(*
SPDX-FileCopyrightText: © 2026 Oleksandr Tiutyk <trofimich@gmail.com>
SPDX-License-Identifier: MIT
License: https://opensource.org/license/mit
*)

(*!
<summary>
Defines the contract for an activity that executes an asynchronous task from TwinCAT.OpenFramework.Tasks.
</summary>
<description>
Starts the task on entry, cyclically executes it while RUNNING, translates stop reasons (WORK_DONE to
completion, INTERNAL_ABORT or EXTERNAL_CANCEL to halted, FAILURE to exception) and propagates cancellation
requests to the task. While suspending, the task keeps executing until it stops. A task failure during
stopping is still an activity failure; work completion completes the activity rather than reporting a pause.
Persistent task bindings distinguish a workflow-owned configuration from an external key.
</description>
*)

INTERFACE IInvokeTaskActivity EXTENDS IActivity

(*!
<summary>Reports whether the task activity has been configured.</summary>
*)
{attribute 'monitoring' := 'call'}
PROPERTY Configured : BOOL
GET
END_GET
END_PROPERTY

(*!
<summary>Configures the task to be executed.</summary>
<description>
Requires a nonzero task instance and PASSIVE_READY. The task is borrowed until stopping and reset finish.
This execution-only binding clears any previously configured persistence role.
Rejected configuration preserves the previous dependency; active task replacement is not supported.
</description>
<param name="task">The task instance to execute.</param>
*)
METHOD Configure
VAR_INPUT
	task : TOF_Tasks.ITask;
END_VAR
END_METHOD

(*!
<summary>Returns the configured task instance, or 0 before configuration.</summary>
*)
{attribute 'monitoring' := 'call'}
PROPERTY Task : TOF_Tasks.ITask
GET
END_GET
END_PROPERTY

(*!
<summary>Adopts a fresh workflow-owned task.</summary>
<description>Requires a ready node in a workflow and a dynamic serializable instance available for exclusive transfer.
The workflow owns it on success. A duplicate in the same workflow raises before changing this node.</description>
*)
METHOD ConfigureEmbeddedTask
VAR_INPUT
	task : TOF_Tasks.ITask;
END_VAR
END_METHOD

(*!
<summary>Binds an externally owned task.</summary>
<description>Requires a live dependency and a nonempty stable key. Several nodes may borrow the same external instance.
The provider keeps it alive. Rejection preserves the previous binding.</description>
*)
METHOD ConfigureExternalTask
VAR_INPUT
	task : TOF_Tasks.ITask;
	key : STRING;
END_VAR
END_METHOD

END_INTERFACE

(* stored: Version 1.1.0.1
   Itf IInvokeTaskActivity: Id {4aac828c-d9ae-42b7-9869-9d06d2ade0db}
   Property Configured: Id {63c9557d-c850-4108-9577-a1cd7c46f917}
   Get Get: Id {39040bea-bdba-45ec-b518-391fda404504}
   Method Configure: Id {50813f6f-26e0-49ce-b6ea-95a18a7ae48d}
   Property Task: Id {6398fb34-b12e-4a05-96cb-c420effe02dc}
   Get Get: Id {3dd712d4-b118-4b87-9656-e8027540988b}
   Method ConfigureEmbeddedTask: Id {4b89e2a9-7271-45ac-b6a7-dfc699ec582e}
   Method ConfigureExternalTask: Id {2ae75d5e-5053-4578-bc2c-d98acda784e7} *)
